Staubli VAL3: DataBase6.pjx

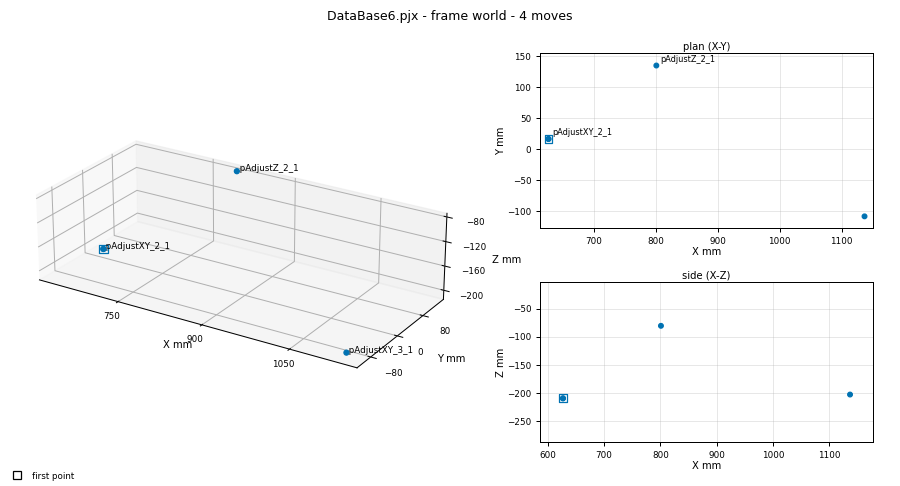
[picture p0: tool path of DataBase6.pjx in frame world, 4 of 24 moves have a stored position in this frame; points joined in program order, loops and branches not executed]
--- DataBase6.pjx ---
Parameters version=s8.10.5Cs9_BS2172 stackSize=5000 millimeterUnit=true
Program file=changeBckColorLabel.pgx
Program file=CheckPosEqual.pgx
Program file=CheckTraj.pgx
Program file=hmiAlert.pgx
Program file=hmiClose.pgx
Program file=hmiConfirm.pgx
Program file=initButton.pgx
Program file=initCheckBox.pgx
Program file=initCombo.pgx
Program file=initContainer.pgx
Program file=initImage.pgx
Program file=initLabel.pgx
Program file=initList.pgx
Program file=initText.pgx
Program file=ListMove.pgx
Program file=moveTarget.pgx
Program file=refreshCheckBox.pgx
Program file=refreshInfo.pgx
Program file=refreshJogMode.pgx
Program file=refreshLanguage.pgx
Program file=refreshQuit.pgx
Program file=updateBtn.pgx
Program file=updateCurrentPos.pgx
Program file=updateInfo.pgx
Program file=updateStr.pgx
Program file=updateTeachPos.pgx
Program file=updateTool.pgx
Data file=DataBase6.dtx
Type name=utButton path=Disk://SmartTCP_CS9/userType/utButton/utButton.pjx
Type name=utCombo path=Disk://SmartTCP_CS9/userType/utCombo/utCombo.pjx
Type name=utContainer path=Disk://SmartTCP_CS9/userType/utContainer/utContainer.pjx
Type name=utImage path=Disk://SmartTCP_CS9/userType/utImage/utImage.pjx
Type name=utLabel path=Disk://SmartTCP_CS9/userType/utLabel/utLabel.pjx
Type name=utList path=Disk://SmartTCP_CS9/userType/utList/utList.pjx
Type name=utText path=Disk://SmartTCP_CS9/userType/utText/utText.pjx
Type name=utTool path=Disk://SmartTCP_CS9/userType/CurrentTool/CurrentTool.pjx

--- DataBase6.dtx ---
public bool bAdjustXY_2_1
public bool bAdjustXY_2_2
public bool bAdjustXY_3_1 = true
public bool bAdjustXY_3_2
public bool bAdjustXY_3_3
public bool bAdjustZ_2_1
public bool bAdjustZ_2_2
public bool bRefresh
public bool bShowJpos
public bool bTeach1 = true
public bool bTeach2 = true
public bool bTeach3 = true
public bool bTeach4 = true
public bool bTeach5
public bool bTeach6
public bool bTeach7
public configRx cConfigSame
public jointRx jAdjustXY_2_1 = {j1=-16.183269, j2=38.957753, j3=100.316368, j4=-129.114182, j5=-108.350352, j6=119.768787}
public jointRx jAdjustXY_2_2 = {j1=-1.561355, j2=34.918272, j3=108.359583, j4=4.917658, j5=-45.199139, j6=85.851346}
public jointRx jAdjustXY_3_1 = {j1=-3.669078, j2=79.701484, j3=49.960672, j4=-7.150792, j5=-35.705417, j6=0.438345}
public jointRx jAdjustXY_3_2 = {j1=19.311169, j2=31.651038, j3=96.790022, j4=84.972086, j5=-76.120044, j6=-139.481694}
public jointRx jAdjustXY_3_3 = {j1=-8.0743577, j2=28.197132, j3=102.272309, j4=-81.334861, j5=-72.794375, j6=-38.960837}
public jointRx jAdjustZ_2_1 = {j1=-3.131112, j2=22.744756, j3=109.0021499, j4=-60.332518, j5=-50.316307, j6=-43.896559}
public jointRx jAdjustZ_2_2 = {j1=-2.340422, j2=42.111372, j3=73.598194, j4=-131.223935, j5=-58.0136019, j6=54.580916}
public jointRx jPosUp
public jointRx jTeach1 = {j1=-3.262771, j2=80.686005, j3=48.0245313, j4=-5.241959, j5=-34.659761, j6=-0.975952}
public jointRx jTeach2 = {j1=-19.636965, j2=85.65368, j3=36.984002, j4=-73.452565, j5=-58.969735, j6=48.957256}
public jointRx jTeach3 = {j1=-1.55114, j2=76.827557, j3=47.134956, j4=16.464605, j5=-15.27397, j6=-40.655038}
public jointRx jTeach4 = {j1=-17.080521, j2=74.155029, j3=36.22097, j4=-118.227611, j5=-47.305779, j6=77.298675}
public jointRx jTeach5
public jointRx jTeach6
public jointRx jTeach7
public mdesc mSlow = {tmax=30, blend=cartesian, leave=0, reach=0}
public mdesc mSpeed_C_blend = {tmax=250, blend=cartesian, leave=0, reach=0}
public mdesc mSpeed_J_blend = {tmax=250, leave=5, reach=5}
public num nBtnItem = 84
public num nClock = 2824.0430321
public num nJogMode = 3
public num nStep0 = 10
public num nStep1 = 11
public num nStep2 = 10
public num nStep3 = 10
public pointRx _pA = {x=1117.817118, y=-89.293345, z=-202.363241, rx=-10.624966, ry=-1.192114, rz=0.674598, shoulder=lefty, elbow=epositive, wrist=wnegative, fatherId=world[0]}
public pointRx _pB = {x=1117.817118, y=-89.293345, z=-202.363241, rx=-2.379148e-15, ry=-1.630783e-17, rz=0.785453, shoulder=lefty, elbow=epositive, wrist=wnegative, fatherId=world[0]}
public pointRx pAdjustXY_2_1 = {x=626.939641, y=16.338855, z=-209.0757962, rx=-0.0000222143, ry=-179.999993, rz=-65.676001, fatherId=world[0]}
public pointRx pAdjustXY_2_2 = {x=857.150616, y=17.401338, z=-208.896815, rx=0.563604, ry=179.453681, rz=42.932806, fatherId=world[0]}
public pointRx pAdjustXY_3_1 = {x=1137.120036, y=-108.57736, z=-202.363161, rx=-0.000297926, ry=0.0000749283, rz=0.78474, shoulder=lefty, elbow=epositive, wrist=wnegative, fatherId=world[0]}
public pointRx pAdjustXY_3_2 = {x=792.594964, y=137.906318, z=-83.726812, rx=0.000088778, ry=179.999738, rz=59.999161, fatherId=world[0]}
public pointRx pAdjustXY_3_3 = {x=785.088371, y=121.389516, z=-83.726812, rx=-0.0000815881, ry=179.99994, rz=-59.999155, fatherId=world[0]}
public pointRx pAdjustZ_2_1 = {x=801.0716396, y=134.899289, z=-80.213051, rx=0.000821012, ry=-179.999765, rz=54.0764076, fatherId=world[0]}
public pointRx pAdjustZ_2_2 = {x=803.315807, y=134.665532, z=-81.371357, rx=0.00172102, ry=-119.999854, rz=54.0779154, fatherId=world[0]}
public pointRx pPosUp = {fatherId=world[0]}
public pointRx pTeach1 = {x=902.313951, y=3.846514, z=-204.254691, rx=-3.799862, ry=94.166562, rz=-1.264999, shoulder=lefty, elbow=epositive, wrist=wnegative, fatherId=world[0]}
public pointRx pTeach2 = {x=880.988773, y=-174.046221, z=-204.254614, rx=82.917358, ry=126.0156651, rz=-89.336459, shoulder=lefty, elbow=epositive, wrist=wnegative, fatherId=world[0]}
public pointRx pTeach3 = {x=911.255756, y=17.873242, z=-173.514595, rx=-16.906456, ry=110.136729, rz=-8.300176, shoulder=lefty, elbow=epositive, wrist=wnegative, fatherId=world[0]}
public pointRx pTeach4 = {x=902.345529, y=-157.209226, z=-88.133434, rx=39.778546, ry=136.990182, rz=-66.473252, shoulder=lefty, elbow=epositive, wrist=wnegative, fatherId=world[0]}
public pointRx pTeach5 = {x=801.894474, y=154.0183518, z=-79.262494, rx=-180, ry=4.770832e-15, rz=180, fatherId=world[0]}
public pointRx pTeach6 = {x=841.843725, y=153.955505, z=-79.296104, rx=-0.00011003, ry=-179.998347, rz=0.00487542, fatherId=world[0]}
public pointRx pTeach7 = {x=841.843706, y=127.954954, z=-79.296104, rx=-0.00022766, ry=-179.998282, rz=0.00522033, fatherId=world[0]}
string sAlertCN{}
  [Align] = "请按Move/Hold键对齐"
  [CantGoBack] = "不可重置!请首先记录第1点!"
  [CantMove1] = "不可到达!请重新记录第1点!"
  [CantMove2] = "不可到达!请重新记录这个点!"
  [CantSwitchTool2] = "不能切换tTool2!请先标定tTool1!"
  [CantSwitchTool3] = "不能切换tTool3!请先标定tTool2!"
  [CompleteAlign] = "对齐完成"
  [CompleteGoBack] = "重置完成"
  [CompleteMove] = "移动完成"
  [DeviationIsTooLarge] = "偏差过大!请重新记录点!"
  [Fifth] = "第5点记录完成"
  [First] = "第1点记录完成"
  [Fourth] = "第4点记录完成"
  [GoBack] = "请按Move/Hold键重置"
  [Move] = "请按Move/Hold键移动"
  [OffsetDone] = "偏差设置完成"
  [Quit] = "您是否决定退出TCP标定应用程序？"
  [SaveInTool1] = "工具参数保存在tTool1"
  [SaveInTool2] = "工具参数保存在tTool2"
  [SaveInTool3] = "工具参数保存在tTool3"
  [Second] = "第2点记录完成"
  [Seventh] = "第7点记录完成"
  [Sixth] = "第6点记录完成"
  [SwitchTool1] = "当前工具已经切换为tTool1!"
  [SwitchTool2] = "当前工具已经切换为tTool2!"
  [SwitchTool3] = "当前工具已经切换为tTool3!"
  [Third] = "第3点记录完成"
  [Version] = "版本: V2.1 日期: 2020.10.12"
string sAlertEN{}
  [Align] = "Press Move/Hold Button To Align"
  [CantGoBack] = "Can't Go back!First record 1st point!"
  [CantMove1] = "Can't Reach!Re-record 1st point!"
  [CantMove2] = "Can't Reach!Re-record this point!"
  [CantSwitchTool2] = "Can't switch to tTool2!Please first calibrate tTool1!"
  [CantSwitchTool3] = "Can't switch to tTool3!Please first calibrate tTool2!"
  [CompleteAlign] = "Alignment has been completed"
  [CompleteGoBack] = "Go back has been completed"
  [CompleteMove] = "Movement has been completed"
  [DeviationIsTooLarge] = "Deviation is too large!Re-record points!"
  [Fifth] = "The 5th point has been recorded"
  [First] = "The 1st point has been recorded"
  [Fourth] = "The 4th point has been recorded"
  [GoBack] = "Press Move/Hold Button to Go back"
  [Move] = "Press Move/Hold Button to Move"
  [OffsetDone] = "Tool deviation has been enabled"
  [Quit] = "Are you sure to quit the tcp calibration application?"
  [SaveInTool1] = "Tool parameters are saved in tTool1"
  [SaveInTool2] = "Tool parameters are saved in tTool2"
  [SaveInTool3] = "Tool parameters are saved in tTool3"
  [Second] = "The 2nd point has been recorded"
  [Seventh] = "The 7th point has been recorded"
  [Sixth] = "The 6th point has been recorded"
  [SwitchTool1] = "The current tool has been switched to tTool1!"
  [SwitchTool2] = "The current tool has been switched to tTool2!"
  [SwitchTool3] = "The current tool has been switched to tTool3!"
  [Third] = "The 3rd point has been recorded"
  [Version] = "Version: V2.1 Date: October 12, 2020"
public string sCbxLanguage = "中文"
public string sCbxMounting = "置顶"
string sHmiCN[200]
  [2] = "语言："
  [3] = "安装："
  [4] = "史陶比尔工具标定 - SmartTCP"
  [7] = "机型："
  [8] = "4轴"
  [9] = "6轴"
  [10] = "工具："
  [11] = "3点标定"
  [12] = "4点标定"
  [13] = "7点标定"
  [14] = "2点180°"
  [15] = "3点120°"
  [16] = "标定工具"
  [17] = "修正工具XY"
  [18] = "修正工具Z"
  [19] = "测试工具"
  [20] = "工具切换："
  [21] = "工具补偿："
  [31] = "点位：P1"
  [32] = "点位：P2"
  [33] = "点位：P3"
  [34] = "点位：P4"
  [35] = "点位：P5"
  [36] = "点位：P6"
  [37] = "点位：P7"
  [41] = "步骤：1/2"
  [42] = "步骤：2/2"
  [43] = "步骤：1/3"
  [44] = "步骤：2/3"
  [45] = "步骤：3/3"
  [46] = "步骤：1/4"
  [47] = "步骤：2/4"
  [48] = "步骤：3/4"
  [49] = "步骤：4/4"
  [50] = "步骤：1/7"
  [51] = "步骤：2/7"
  [52] = "步骤：3/7"
  [53] = "步骤：4/7"
  [54] = "步骤：5/7"
  [55] = "步骤：6/7"
  [56] = "步骤：7/7"
  [80] = "对齐,记录,移动,Null,Null,Null,返回,继续"
  [81] = "Null,记录,移动,Null,Null,Null,返回,继续"
  [82] = "Null,记录,移动,Null,Null,计算,返回,完成"
  [83] = "Null,Null,Null,Null,Null,Null,Null,退出"
  [84] = "对齐,记录,移动,切换,Null,Null,返回,继续"
  [85] = "重置,记录,移动,RZ+,RZ-,计算,返回,完成"
  [86] = "重置,记录,移动,RZ+,Null,Null,返回,继续"
  [87] = "重置,记录,移动,RZ-,Null,计算,返回,完成"
  [88] = "重置,记录,移动,RX+,RY+,计算,返回,完成"
  [89] = "对齐,Null,Null,Null,Null,Null,Null,完成"
  [100] = "适配TX2/TS2机器人的工具标定应用程序"
  [101] = "操作提醒："
  [102] = "工具垂直姿态对准尖点并记录"
  [103] = "工具任意姿态对准尖点并记录"
  [104] = "按计算按钮获取TCP值"
  [105] = "按记录按钮保存当前位置"
  [106] = "按记录按钮保存当前位置（坐标系原点）"
  [107] = "按记录按钮保存当前位置（坐标系OX方向）"
  [108] = "按记录按钮保存当前位置（坐标系OXY平面）"
  [109] = "保持当前姿态沿X方向移动"
  [110] = "保持当前姿态沿Y方向移动"
  [111] = "确保TCP(RZ) 可以反向旋转180°"
  [112] = "按RZ+(RZ-)与Move/Hold按钮旋转TCP 180°"
  [113] = "旋转TCP(RZ)接近一侧极限"
  [114] = "旋转TCP(RZ)接近中间位置"
  [115] = "确保TCP(RZ) 可以旋转±60°"
  [116] = "按RZ+与Move/Hold按钮旋转TCP +60°"
  [117] = "按RZ-与Move/Hold按钮旋转TCP -60°"
  [118] = "确保TCP(RY)或 TCP(RX)可以旋转+60°"
  [119] = "按RX+(RY+)与Move/Hold按钮旋转TCP +60°"
  [120] = "工具当前姿态对准尖点并记录"
  [121] = "最大可旋转角度只有:"
  [125] = "对齐适用于用户工具与法兰轴向为90°的情况"
string sHmiEN[200]
  [2] = "Language："
  [3] = "Mounting："
  [4] = "Stäubli Tool Calibration - SmartTCP"
  [7] = "ArmType："
  [8] = "4Axis"
  [9] = "6Axis"
  [10] = "Tool："
  [11] = "3Points"
  [12] = "4Points"
  [13] = "7Points"
  [14] = "2Points180°"
  [15] = "3Points120°"
  [16] = "Calibration tool"
  [17] = "Correction tool XY"
  [18] = "Correction tool Z"
  [19] = "Verification tool"
  [20] = "Tool Switch："
  [21] = "Tool Offset："
  [31] = "Point：P1"
  [32] = "Point：P2"
  [33] = "Point：P3"
  [34] = "Point：P4"
  [35] = "Point：P5"
  [36] = "Point：P6"
  [37] = "Point：P7"
  [41] = "Step：1/2"
  [42] = "Step：2/2"
  [43] = "Step：1/3"
  [44] = "Step：2/3"
  [45] = "Step：3/3"
  [46] = "Step：1/4"
  [47] = "Step：2/4"
  [48] = "Step：3/4"
  [49] = "Step：4/4"
  [50] = "Step：1/7"
  [51] = "Step：2/7"
  [52] = "Step：3/7"
  [53] = "Step：4/7"
  [54] = "Step：5/7"
  [55] = "Step：6/7"
  [56] = "Step：7/7"
  [80] = "Align,Here,Move,Null,Null,Null,Prev.,Next"
  [81] = "Null,Here,Move,Null,Null,Null,Prev.,Next"
  [82] = "Null,Here,Move,Null,Null,Calc.,Prev.,Done"
  [83] = "Null,Null,Null,Null,Null,Null,Null,Quit"
  [84] = "Align,Here,Move,Chg.,Null,Null,Prev.,Next"
  [85] = "Reset,Here,Move,RZ+,RZ-,Calc.,Prev.,Done"
  [86] = "Reset,Here,Move,RZ+,Null,Null,Prev.,Next"
  [87] = "Reset,Here,Move,RZ-,Null,Calc.,Prev.,Done"
  [88] = "Reset,Here,Move,RX+,RY+,Calc.,Prev.,Done"
  [89] = "Align,Null,Null,Null,Null,Null,Null,Done"
  [100] = "TCP calibration application for TX2/TS2 robot"
  [101] = "Operation reminder："
  [102] = "Touch to reference pointer in vertical attitude"
  [103] = "Touch to reference pointer in any attitude"
  [104] = "Press Calc. button to get the TCP value"
  [105] = "Press Here button to save the position"
  [106] = "Press Here button to save the position (Frame Origin)"
  [107] = "Press Here button to save the position (Frame Axis OX)"
  [108] = "Press Here button to save the position (Frame Plane OXY)"
  [109] = "Keep the current attitude moving in X direction"
  [110] = "Keep the current attitude moving in Y direction"
  [111] = "Ensure that the TCP(RZ) reverse can be rotated 180°"
  [112] = "Press the RZ+(RZ-) & Move/Hold to rotate TCP 180°"
  [113] = "Rotate TCP (RZ) close to one side limit"
  [114] = "Rotate TCP (RZ) close to middle position"
  [115] = "Ensure that the TCP(RZ) can be rotated ±60°"
  [116] = "Press the RZ+ & Move/Hold to rotate TCP +60°"
  [117] = "Press the RZ- & Move/Hold to rotate TCP -60°"
  [118] = "Ensure that the TCP(RX) or TCP(RY) can be rotated +60°"
  [119] = "Press the RX+(RY+) & Move/Hold to rotate TCP +60°"
  [120] = "Touch to reference pointer in current attitude"
  [121] = "The maximum rotation angle is only:"
  [125] = "Alignment can be used when the tool and flange are 90°"
public string sLanguage = "chinese"
public string sLanguageM = "chinese"
public string sMounting = "Ceiling"
public tool tCurrentTool = {x=-7.678916, y=-111.709078, z=238.876751, rx=-50.589367, ry=-96.556923, rz=-50.497076, fatherId=flange[0], ioLink=FastIO\fOut0}
public tool tFlange = {fatherId=flange[0]}
public tool tTool1 = {x=-7.678916, y=-111.709078, z=238.876751, rx=-50.589367, ry=-96.556923, rz=-50.497076, fatherId=flange[0], ioLink=FastIO\fOut0}
public tool tTool2 = {x=12.349519, y=146.187295, z=111.945303, rx=-81.862508, ry=5.143902, rz=-177.300649, fatherId=flange[0], ioLink=FastIO\fOut0}
public tool tTool3 = {x=11, y=22, z=33, rx=20, ry=30, rz=40, fatherId=flange[0], ioLink=FastIO\fOut0}
public trsf trOffset = {z=10}
public trsf trOffsetM = {x=11, y=22, z=33, rx=44, ry=55, rz=66}
public utButton utBtn_Bottom[8]
  [0]
    utAppearance Appearance
      [0]
        bool bVisibility = true
        string sBackgroundColour = "#FFFFFF"
        string sBackgroundImage
        string sColour
    utBorder Border
      [0]
        string sBorderColour
    utCommon Common
      [0]
        bool bDisabled
        string sID = "bottom_btn0"
        string sPage = "Disk://SmartTCP_CS9/tx2/interface/Page_Main"
        string sText = "对齐"
    utData Data
      [0]
        bool bStatus
        num nVal
    utEvents Events
      [0]
        bool bClick
        bool bMouseDown
        bool bMouseUp
    utText Text
      [0]
        num nFontSize
        string sFontFamily
        string sFontStyle
        string sFontWeight
        string sTextAlignment
  [1]
    utAppearance Appearance
      [0]
        bool bVisibility = true
        string sBackgroundColour = "#FFFFFF"
        string sBackgroundImage
        string sColour
    utBorder Border
      [0]
        string sBorderColour
    utCommon Common
      [0]
        bool bDisabled
        string sID = "bottom_btn1"
        string sPage = "Disk://SmartTCP_CS9/tx2/interface/Page_Main"
        string sText = "记录"
    utData Data
      [0]
        bool bStatus
        num nVal
    utEvents Events
      [0]
        bool bClick
        bool bMouseDown
        bool bMouseUp
    utText Text
      [0]
        num nFontSize
        string sFontFamily
        string sFontStyle
        string sFontWeight
        string sTextAlignment
  [2]
    utAppearance Appearance
      [0]
        bool bVisibility = true
        string sBackgroundColour = "#FFFFFF"
        string sBackgroundImage
        string sColour
    utBorder Border
      [0]
        string sBorderColour
    utCommon Common
      [0]
        bool bDisabled
        string sID = "bottom_btn2"
        string sPage = "Disk://SmartTCP_CS9/tx2/interface/Page_Main"
        string sText = "移动"
    utData Data
      [0]
        bool bStatus
        num nVal
    utEvents Events
      [0]
        bool bClick
        bool bMouseDown
        bool bMouseUp
    utText Text
      [0]
        num nFontSize
        string sFontFamily
        string sFontStyle
        string sFontWeight
        string sTextAlignment
  [3]
    utAppearance Appearance
      [0]
        bool bVisibility = true
        string sBackgroundColour = "#FFFFFF"
        string sBackgroundImage
        string sColour
    utBorder Border
      [0]
        string sBorderColour
    utCommon Common
      [0]
        bool bDisabled
        string sID = "bottom_btn3"
        string sPage = "Disk://SmartTCP_CS9/tx2/interface/Page_Main"
        string sText = "切换"
    utData Data
      [0]
        bool bStatus
        num nVal
    utEvents Events
      [0]
        bool bClick
        bool bMouseDown
        bool bMouseUp
    utText Text
      [0]
        num nFontSize
        string sFontFamily
        string sFontStyle
        string sFontWeight
        string sTextAlignment
  [4]
    utAppearance Appearance
      [0]
        bool bVisibility
        string sBackgroundColour = "#FFFFFF"
        string sBackgroundImage
        string sColour
    utBorder Border
      [0]
        string sBorderColour
    utCommon Common
      [0]
        bool bDisabled
        string sID = "bottom_btn4"
        string sPage = "Disk://SmartTCP_CS9/tx2/interface/Page_Main"
        string sText
    utData Data
      [0]
        bool bStatus
        num nVal
    utEvents Events
      [0]
        bool bClick
        bool bMouseDown
        bool bMouseUp
    utText Text
      [0]
        num nFontSize
        string sFontFamily
        string sFontStyle
        string sFontWeight
        string sTextAlignment
  [5]
    utAppearance Appearance
      [0]
        bool bVisibility
        string sBackgroundColour = "#FFFFFF"
        string sBackgroundImage
        string sColour
    utBorder Border
      [0]
        string sBorderColour
    utCommon Common
      [0]
        bool bDisabled
        string sID = "bottom_btn5"
        string sPage = "Disk://SmartTCP_CS9/tx2/interface/Page_Main"
        string sText
    utData Data
      [0]
        bool bStatus
        num nVal
    utEvents Events
      [0]
        bool bClick
        bool bMouseDown
        bool bMouseUp
    utText Text
      [0]
        num nFontSize
        string sFontFamily
        string sFontStyle
        string sFontWeight
        string sTextAlignment
  [6]
    utAppearance Appearance
      [0]
        bool bVisibility = true
        string sBackgroundColour = "#FFFFFF"
        string sBackgroundImage
        string sColour
    utBorder Border
      [0]
        string sBorderColour
    utCommon Common
      [0]
        bool bDisabled
        string sID = "bottom_btn6"
        string sPage = "Disk://SmartTCP_CS9/tx2/interface/Page_Main"
        string sText = "返回"
    utData Data
      [0]
        bool bStatus
        num nVal
    utEvents Events
      [0]
        bool bClick
        bool bMouseDown
        bool bMouseUp
    utText Text
      [0]
        num nFontSize
        string sFontFamily
        string sFontStyle
        string sFontWeight
        string sTextAlignment
  [7]
    utAppearance Appearance
      [0]
        bool bVisibility = true
        string sBackgroundColour = "#FFFFFF"
        string sBackgroundImage
        string sColour
    utBorder Border
      [0]
        string sBorderColour
    utCommon Common
      [0]
        bool bDisabled
        string sID = "bottom_btn7"
        string sPage = "Disk://SmartTCP_CS9/tx2/interface/Page_Main"
        string sText = "继续"
    utData Data
      [0]
        bool bStatus
        num nVal
    utEvents Events
      [0]
        bool bClick
        bool bMouseDown
        bool bMouseUp
    utText Text
      [0]
        num nFontSize
        string sFontFamily
        string sFontStyle
        string sFontWeight
        string sTextAlignment
public utButton utBtn_No
  [0]
    utAppearance Appearance
      [0]
        bool bVisibility = true
        string sBackgroundColour = "#FFFFFF"
        string sBackgroundImage
        string sColour
    utBorder Border
      [0]
        string sBorderColour
    utCommon Common
      [0]
        bool bDisabled
        string sID = "btn_No"
        string sPage = "Disk://SmartTCP_CS9/tx2/interface/Page_Container_Confirm"
        string sText = "No"
    utData Data
      [0]
        bool bStatus
        num nVal
    utEvents Events
      [0]
        bool bClick
        bool bMouseDown
        bool bMouseUp
    utText Text
      [0]
        num nFontSize
        string sFontFamily
        string sFontStyle
        string sFontWeight
        string sTextAlignment
public utButton utBtn_OK
  [0]
    utAppearance Appearance
      [0]
        bool bVisibility = true
        string sBackgroundColour = "#FFFFFF"
        string sBackgroundImage
        string sColour
    utBorder Border
      [0]
        string sBorderColour
    utCommon Common
      [0]
        bool bDisabled
        string sID = "btn_OK"
        string sPage = "Disk://SmartTCP_CS9/tx2/interface/Page_Container_Alert"
        string sText = "OK"
    utData Data
      [0]
        bool bStatus
        num nVal
    utEvents Events
      [0]
        bool bClick
        bool bMouseDown
        bool bMouseUp
    utText Text
      [0]
        num nFontSize
        string sFontFamily
        string sFontStyle
        string sFontWeight
        string sTextAlignment
public utButton utBtn_Step[4]
  [0]
    utAppearance Appearance
      [0]
        bool bVisibility = true
        string sBackgroundColour = "#FFFFFF"
        string sBackgroundImage
        string sColour
    utBorder Border
      [0]
        string sBorderColour
    utCommon Common
      [0]
        bool bDisabled
        string sID = "step_btn0"
        string sPage = "Disk://SmartTCP_CS9/tx2/interface/Page_Container_Main"
        string sText = "标定工具"
    utData Data
      [0]
        bool bStatus
        num nVal = 16
    utEvents Events
      [0]
        bool bClick
        bool bMouseDown
        bool bMouseUp
    utText Text
      [0]
        num nFontSize
        string sFontFamily
        string sFontStyle
        string sFontWeight
        string sTextAlignment
  [1]
    utAppearance Appearance
      [0]
        bool bVisibility = true
        string sBackgroundColour = "#FFFFFF"
        string sBackgroundImage
        string sColour
    utBorder Border
      [0]
        string sBorderColour
    utCommon Common
      [0]
        bool bDisabled
        string sID = "step_btn1"
        string sPage = "Disk://SmartTCP_CS9/tx2/interface/Page_Container_Main"
        string sText = "修正工具XY"
    utData Data
      [0]
        bool bStatus
        num nVal = 17
    utEvents Events
      [0]
        bool bClick = true
        bool bMouseDown
        bool bMouseUp
    utText Text
      [0]
        num nFontSize
        string sFontFamily
        string sFontStyle
        string sFontWeight
        string sTextAlignment
  [2]
    utAppearance Appearance
      [0]
        bool bVisibility = true
        string sBackgroundColour = "#FFFFFF"
        string sBackgroundImage
        string sColour
    utBorder Border
      [0]
        string sBorderColour
    utCommon Common
      [0]
        bool bDisabled
        string sID = "step_btn2"
        string sPage = "Disk://SmartTCP_CS9/tx2/interface/Page_Container_Main"
        string sText = "修正工具Z"
    utData Data
      [0]
        bool bStatus
        num nVal = 18
    utEvents Events
      [0]
        bool bClick
        bool bMouseDown
        bool bMouseUp
    utText Text
      [0]
        num nFontSize
        string sFontFamily
        string sFontStyle
        string sFontWeight
        string sTextAlignment
  [3]
    utAppearance Appearance
      [0]
        bool bVisibility = true
        string sBackgroundColour = "#FFFFFF"
        string sBackgroundImage
        string sColour
    utBorder Border
      [0]
        string sBorderColour
    utCommon Common
      [0]
        bool bDisabled
        string sID = "step_btn3"
        string sPage = "Disk://SmartTCP_CS9/tx2/interface/Page_Container_Main"
        string sText = "测试工具"
    utData Data
      [0]
        bool bStatus
        num nVal = 19
    utEvents Events
      [0]
        bool bClick
        bool bMouseDown
        bool bMouseUp
    utText Text
      [0]
        num nFontSize
        string sFontFamily
        string sFontStyle
        string sFontWeight
        string sTextAlignment
public utButton utBtn_Yes
  [0]
    utAppearance Appearance
      [0]
        bool bVisibility = true
        string sBackgroundColour = "#FFFFFF"
        string sBackgroundImage
        string sColour
    utBorder Border
      [0]
        string sBorderColour
    utCommon Common
      [0]
        bool bDisabled
        string sID = "btn_Yes"
        string sPage = "Disk://SmartTCP_CS9/tx2/interface/Page_Container_Confirm"
        string sText = "Yes"
    utData Data
      [0]
        bool bStatus
        num nVal
    utEvents Events
      [0]
        bool bClick
        bool bMouseDown
        bool bMouseUp
    utText Text
      [0]
        num nFontSize
        string sFontFamily
        string sFontStyle
        string sFontWeight
        string sTextAlignment
public utCombo utCbx_Language_Data
  [0]
    utAppearance Appearance
      [0]
        bool bVisibility
        string sBackgroundColour
        string sColour
    utBorder Border
      [0]
        string sBorderColour
        string sBorderStyle
        string sBorderWidth
    utCommon Common
      [0]
        bool bDisabled
        string sID = "cbx_Language_D"
        string sItem[2]
          [0] = "中文"
          [1] = "英文"
        string sOption{}
        string sPage = "Disk://SmartTCP_CS9/tx2/interface/Page_Main"
        string sValue = "中文"
    utData Data
      [0]
        bool bStatus
        num nVal
    utText Text
      [0]
        num nFontSize
        string sFontFamily
        string sFontStyle
public utCombo utCbx_Mounting_Data
  [0]
    utAppearance Appearance
      [0]
        bool bVisibility
        string sBackgroundColour
        string sColour
    utBorder Border
      [0]
        string sBorderColour
        string sBorderStyle
        string sBorderWidth
    utCommon Common
      [0]
        bool bDisabled
        string sID = "cbx_Mounting_D"
        string sItem[2]
          [0] = "置地"
          [1] = "置顶"
        string sOption{}
        string sPage = "Disk://SmartTCP_CS9/tx2/interface/Page_Main"
        string sValue = "置顶"
    utData Data
      [0]
        bool bStatus
        num nVal
    utText Text
      [0]
        num nFontSize
        string sFontFamily
        string sFontStyle
public utContainer utCtn_Function
  [0]
    utAppearance Appearance
      [0]
        bool bVisibility = true
    utCommon Common
      [0]
        string sID = "ctn_Function"
        string sPage = "Disk://SmartTCP_CS9/tx2/interface/Page_Main"
        string sSource = "Page_Container_Teach.html"
public utContainer utCtn_Message
  [0]
    utAppearance Appearance
      [0]
        bool bVisibility
    utCommon Common
      [0]
        string sID = "ctn_Message"
        string sPage = "Disk://SmartTCP_CS9/tx2/interface/Page_Main"
        string sSource = "Page_Container_Alert.html"
public utImage utImg_CheckBox_a[3]
  [0]
    utAppearance Appearance
      [0]
        bool bVisibility
        string sBackgroundColour
    utBorder Border
      [0]
        num nBorderWidth
        string sBorderColour
        string sBorderStyle
    utCommon Common
      [0]
        string sClass = "clickable"
        string sID = "img_CheckBox_a0"
        string sPage = "Disk://SmartTCP_CS9/tx2/interface/Page_Container_Main"
        string sSourceImage = "images/checkbox_unchecked.png"
    utData Data
      [0]
        bool bStatus
        num nVal
        string sSourceImg1 = "images/checkbox_checked.png"
        string sSourceImg2 = "images/checkbox_unchecked.png"
    utEvents Events
      [0]
        bool bClick
        bool bMouseDown
        bool bMouseUp
  [1]
    utAppearance Appearance
      [0]
        bool bVisibility
        string sBackgroundColour
    utBorder Border
      [0]
        num nBorderWidth
        string sBorderColour
        string sBorderStyle
    utCommon Common
      [0]
        string sClass = "clickable"
        string sID = "img_CheckBox_a1"
        string sPage = "Disk://SmartTCP_CS9/tx2/interface/Page_Container_Main"
        string sSourceImage = "images/checkbox_checked.png"
    utData Data
      [0]
        bool bStatus = true
        num nVal
        string sSourceImg1 = "images/checkbox_checked.png"
        string sSourceImg2 = "images/checkbox_unchecked.png"
    utEvents Events
      [0]
        bool bClick
        bool bMouseDown
        bool bMouseUp
  [2]
    utAppearance Appearance
      [0]
        bool bVisibility
        string sBackgroundColour
    utBorder Border
      [0]
        num nBorderWidth
        string sBorderColour
        string sBorderStyle
    utCommon Common
      [0]
        string sClass = "clickable"
        string sID = "img_CheckBox_a2"
        string sPage = "Disk://SmartTCP_CS9/tx2/interface/Page_Container_Main"
        string sSourceImage = "images/checkbox_unchecked.png"
    utData Data
      [0]
        bool bStatus
        num nVal
        string sSourceImg1 = "images/checkbox_checked.png"
        string sSourceImg2 = "images/checkbox_unchecked.png"
    utEvents Events
      [0]
        bool bClick
        bool bMouseDown
        bool bMouseUp
public utImage utImg_CheckBox_b[2]
  [0]
    utAppearance Appearance
      [0]
        bool bVisibility
        string sBackgroundColour
    utBorder Border
      [0]
        num nBorderWidth
        string sBorderColour
        string sBorderStyle
    utCommon Common
      [0]
        string sClass = "clickable"
        string sID = "img_CheckBox_b0"
        string sPage = "Disk://SmartTCP_CS9/tx2/interface/Page_Container_Main"
        string sSourceImage = "images/checkbox_unchecked.png"
    utData Data
      [0]
        bool bStatus
        num nVal
        string sSourceImg1 = "images/checkbox_checked.png"
        string sSourceImg2 = "images/checkbox_unchecked.png"
    utEvents Events
      [0]
        bool bClick
        bool bMouseDown
        bool bMouseUp
  [1]
    utAppearance Appearance
      [0]
        bool bVisibility
        string sBackgroundColour
    utBorder Border
      [0]
        num nBorderWidth
        string sBorderColour
        string sBorderStyle
    utCommon Common
      [0]
        string sClass = "clickable"
        string sID = "img_CheckBox_b1"
        string sPage = "Disk://SmartTCP_CS9/tx2/interface/Page_Container_Main"
        string sSourceImage = "images/checkbox_checked.png"
    utData Data
      [0]
        bool bStatus = true
        num nVal
        string sSourceImg1 = "images/checkbox_checked.png"
        string sSourceImg2 = "images/checkbox_unchecked.png"
    utEvents Events
      [0]
        bool bClick
        bool bMouseDown
        bool bMouseUp
public utImage utImg_Example
  [0]
    utAppearance Appearance
      [0]
        bool bVisibility = true
        string sBackgroundColour
    utBorder Border
      [0]
        num nBorderWidth
        string sBorderColour
        string sBorderStyle
    utCommon Common
      [0]
        string sClass = "clickable"
        string sID = "img_example"
        string sPage = "Disk://SmartTCP_CS9/tx2/interface/Page_Container_Teach"
        string sSourceImage = "images/6AxisAdjustXY2_1.png"
    utData Data
      [0]
        bool bStatus
        num nVal
        string sSourceImg1
        string sSourceImg2
    utEvents Events
      [0]
        bool bClick
        bool bMouseDown
        bool bMouseUp
public utImage utImg_Info
  [0]
    utAppearance Appearance
      [0]
        bool bVisibility = true
        string sBackgroundColour
    utBorder Border
      [0]
        num nBorderWidth
        string sBorderColour
        string sBorderStyle
    utCommon Common
      [0]
        string sClass = "clickable"
        string sID = "img_info"
        string sPage = "Disk://SmartTCP_CS9/tx2/interface/Page_Main"
        string sSourceImage = "images/info.png"
    utData Data
      [0]
        bool bStatus
        num nVal
        string sSourceImg1 = "images/switch_on.png"
        string sSourceImg2 = "images/switch_off.png"
    utEvents Events
      [0]
        bool bClick
        bool bMouseDown
        bool bMouseUp
public utImage utImg_JogMode[4]
  [0]
    utAppearance Appearance
      [0]
        bool bVisibility = true
        string sBackgroundColour
    utBorder Border
      [0]
        num nBorderWidth
        string sBorderColour = "#000000"
        string sBorderStyle = "Solid"
    utCommon Common
      [0]
        string sClass = "clickable"
        string sID = "img_None"
        string sPage = "Disk://SmartTCP_CS9/tx2/interface/Page_Main"
        string sSourceImage = "images/none.svg"
    utData Data
      [0]
        bool bStatus
        num nVal
        string sSourceImg1
        string sSourceImg2
    utEvents Events
      [0]
        bool bClick
        bool bMouseDown
        bool bMouseUp
  [1]
    utAppearance Appearance
      [0]
        bool bVisibility = true
        string sBackgroundColour
    utBorder Border
      [0]
        num nBorderWidth
        string sBorderColour = "#FFFFFF"
        string sBorderStyle = "None"
    utCommon Common
      [0]
        string sClass = "clickable"
        string sID = "img_Joint"
        string sPage = "Disk://SmartTCP_CS9/tx2/interface/Page_Main"
        string sSourceImage = "images/joint.svg"
    utData Data
      [0]
        bool bStatus
        num nVal
        string sSourceImg1
        string sSourceImg2
    utEvents Events
      [0]
        bool bClick
        bool bMouseDown
        bool bMouseUp
  [2]
    utAppearance Appearance
      [0]
        bool bVisibility = true
        string sBackgroundColour
    utBorder Border
      [0]
        num nBorderWidth
        string sBorderColour = "#FFFFFF"
        string sBorderStyle = "None"
    utCommon Common
      [0]
        string sClass = "clickable"
        string sID = "img_Frame"
        string sPage = "Disk://SmartTCP_CS9/tx2/interface/Page_Main"
        string sSourceImage = "images/frame.svg"
    utData Data
      [0]
        bool bStatus
        num nVal
        string sSourceImg1
        string sSourceImg2
    utEvents Events
      [0]
        bool bClick
        bool bMouseDown
        bool bMouseUp
  [3]
    utAppearance Appearance
      [0]
        bool bVisibility = true
        string sBackgroundColour
    utBorder Border
      [0]
        num nBorderWidth
        string sBorderColour = "#FFFFFF"
        string sBorderStyle = "None"
    utCommon Common
      [0]
        string sClass = "selected"
        string sID = "img_Tool"
        string sPage = "Disk://SmartTCP_CS9/tx2/interface/Page_Main"
        string sSourceImage = "images/tool.svg"
    utData Data
      [0]
        bool bStatus
        num nVal
        string sSourceImg1
        string sSourceImg2
    utEvents Events
      [0]
        bool bClick
        bool bMouseDown
        bool bMouseUp
public utImage utImg_Next
  [0]
    utAppearance Appearance
      [0]
        bool bVisibility = true
        string sBackgroundColour
    utBorder Border
      [0]
        num nBorderWidth
        string sBorderColour
        string sBorderStyle
    utCommon Common
      [0]
        string sClass = "clickable"
        string sID = "img_Next"
        string sPage = "Disk://SmartTCP_CS9/tx2/interface/Page_Container_Test"
        string sSourceImage = "images/navigate-next.svg"
    utData Data
      [0]
        bool bStatus
        num nVal
        string sSourceImg1
        string sSourceImg2
    utEvents Events
      [0]
        bool bClick
        bool bMouseDown
        bool bMouseUp
public utImage utImg_PosSwitch
  [0]
    utAppearance Appearance
      [0]
        bool bVisibility = true
        string sBackgroundColour
    utBorder Border
      [0]
        num nBorderWidth
        string sBorderColour
        string sBorderStyle
    utCommon Common
      [0]
        string sClass = "clickable"
        string sID = "img_PosSwitch"
        string sPage = "Disk://SmartTCP_CS9/tx2/interface/Page_Main"
        string sSourceImage = "images/switch.png"
    utData Data
      [0]
        bool bStatus
        num nVal
        string sSourceImg1
        string sSourceImg2
    utEvents Events
      [0]
        bool bClick
        bool bMouseDown
        bool bMouseUp
public utImage utImg_Previous
  [0]
    utAppearance Appearance
      [0]
        bool bVisibility = true
        string sBackgroundColour
    utBorder Border
      [0]
        num nBorderWidth
        string sBorderColour
        string sBorderStyle
    utCommon Common
      [0]
        string sClass = "clickable"
        string sID = "img_Previous"
        string sPage = "Disk://SmartTCP_CS9/tx2/interface/Page_Container_Test"
        string sSourceImage = "images/navigate-previous.svg"
    utData Data
      [0]
        bool bStatus
        num nVal
        string sSourceImg1
        string sSourceImg2
    utEvents Events
      [0]
        bool bClick
        bool bMouseDown
        bool bMouseUp
public utImage utImg_Switch
  [0]
    utAppearance Appearance
      [0]
        bool bVisibility
        string sBackgroundColour
    utBorder Border
      [0]
        num nBorderWidth
        string sBorderColour
        string sBorderStyle
    utCommon Common
      [0]
        string sClass = "clickable"
        string sID = "img_Switch"
        string sPage = "Disk://SmartTCP_CS9/tx2/interface/Page_Container_Test"
        string sSourceImage = "images/switch_off.png"
    utData Data
      [0]
        bool bStatus
        num nVal
        string sSourceImg1 = "images/switch_on.png"
        string sSourceImg2 = "images/switch_off.png"
    utEvents Events
      [0]
        bool bClick
        bool bMouseDown
        bool bMouseUp
public utLabel utLbl_Axis
  [0]
    utAppearance Appearance
      [0]
        bool bVisibility
        string sBackgroundColour = "#FFFFFF"
        string sColour
    utBorder Border
      [0]
        num nBorderWidth
